Fanuc KAREL source: kf00050.KL

-- PROVISIONAL review KL for V770-1; original PC SHA256 dc6943842294447fd62e46bbde16faa84ccde77ae134d5c3726c594ab87717b8
-- Incomplete behavior may be omitted. Consult companion uncertainty JSON. Do not deploy.
PROGRAM KF00050
%NOLOCKGROUP
VAR
  I : INTEGER
  J : INTEGER
  X : REAL
  Y : REAL
  B : BOOLEAN
  C : BOOLEAN
  TXT : STRING[80]
  TXT2 : STRING[80]
  STATUS : INTEGER
-- UNRESOLVED_DECL AI type=002010
-- UNRESOLVED_DECL BI type=002010
-- UNRESOLVED_DECL P type=000102
-- UNRESOLVED_DECL JP type=000199
-- UNRESOLVED_DECL PF type=000101
-- UNRESOLVED_DECL V1 type=000013
-- UNRESOLVED_DECL V2 type=000013
BEGIN
  -- UNRESOLVED_PC offsets 5-34; opcodes 9D,23,9E,2E,22,7A
  -- UNRESOLVED_PC offsets 39-58; opcodes 21,21,52,23
  -- UNRESOLVED_PC offsets 63-78; opcodes 20,2C,23
  -- UNRESOLVED_PC offsets 83-87; opcodes 7F
END KF00050
